(* PLC project Vn_fbd_set_output, Beckhoff Automation GmbH TwinCAT PLC Control 3.5.13.21 *)
(* stored: creationDateTime 1970-01-01T00:00:00 *)

PROGRAM Vn_fbd_set_output

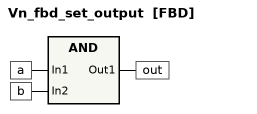
(* FBD diagram, written out as Structured Text *)
IF a AND b THEN out := TRUE; END_IF;
END_PROGRAM
